ABB RAPID module: LongProg_3.mod

%%%
  VERSION:1
  LANGUAGE:ENGLISH
%%%
MODULE MOD_Tmp1

	PROC Prg_Tmp1()

		MoveAbsJ [[500.000000,0.000000,0.000000,0.000000,0.000000,0.000000],[9E+09,9E+09,9E+09,9E+09,9E+09,9E+09]],v500,z1,ToolS \WObj:=FrameS;

	ENDPROC

ENDMODULE
